KUKA KRL program: PgProg.src

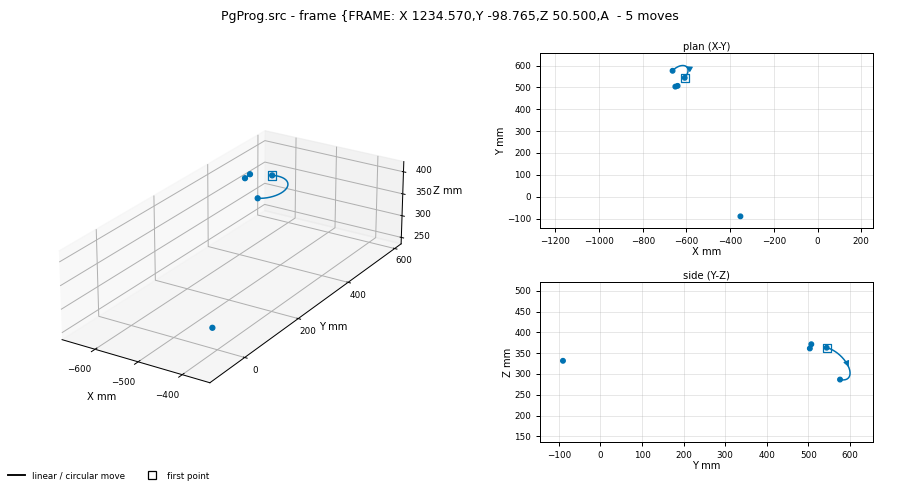
[picture p0: tool path of PgProg.src in frame {FRAME: X 1234.570,Y -98.765,Z 50.500,A , 5 of 9 moves have a stored position in this frame; points joined in program order, loops and branches not executed]
&ACCESS RVP
&REL 1
&PARAM TEMPLATE = C:\KRC\Roboter\Template\vorgabe
&PARAM EDITMASK = *
DEF PgProg ( )


; GLOBAL INTERRUPT DECL 3 WHEN $STOPMESS==TRUE DO IR_STOPM ( )
; INTERRUPT ON 3

;FOLD Initialise and set default speed
BAS (#INITMOV,0)
BAS (#VEL_PTP,100)
BAS (#ACC_PTP,20)
$VEL.CP=0.2
BAS (#TOOL,0)
BAS (#BASE,0)
;ENDFOLD

;;FOLD STARTPOS
;$BWDSTART = FALSE
;PDAT_ACT = PDEFAULT
;BAS(#PTP_DAT)
;FDAT_ACT = {TOOL_NO 0,BASE_NO 0,IPO_FRAME #BASE}
;BAS(#FRAMES)
;;ENDFOLD

$ADVANCE = 5

;FOLD ---- Quickly skip BCO ----
; PTP $AXIS_ACT
;ENDFOLD

;FOLD ---- GO HOME ----
; PTP {A1 0.000, A2 -90.000, A3 90.000, A4 0.000, A5 0.000, A6 0.000, E1 0, E2 0, E3 0, E4 0, E5 0, E6 0}
;ENDFOLD


; Program generated by RoboDK v6.0.7 for KUKA KR 10 R1440-2 on XX/XX/XXXX 18:00:00
; Using nominal kinematics.
; ---- Setting reference (Base) ----
$BASE = {FRAME: X 1234.570,Y -98.765,Z 50.500,A 30.000,B 0.000,C 0.000}
; --------------------------
; ---- Setting tool (TCP) ----
$TOOL = {FRAME: X 10.000,Y 20.000,Z 150.000,A 0.000,B 0.000,C 15.000}
; --------------------------
$VEL.CP = 0.25000
$APO.CPTP = 5
$APO.CDIS = 5.000
PTP {A1 0.00000,A2 -10.00000,A3 20.00000,A4 0.00000,A5 30.00000,A6 0.00000} C_PTP
LIN {X -607.850,Y 543.849,Z 363.215,A 150.000,B 50.000,C -165.000} C_DIS
CIRC {X -602.951,Y 596.788,Z 316.595,A 150.000,B 50.000,C -165.000},{X -663.517,Y 575.988,Z 286.611,A 150.000,B 50.000,C -165.000} C_DIS
PTP {A1 20.00000,A2 -10.00000,A3 20.00000,A4 0.00000,A5 30.00000,A6 0.00000} C_PTP
$ACC.ORI1 = 120.00000
$ACC.ORI2 = 120.00000
$VEL.ORI1 = 60.00000
$VEL.ORI2 = 60.00000
$ACC.CP = 0.80000
$VEL.CP = 0.10000
LIN {X -650.861,Y 503.437,Z 361.399,A 150.000,B 50.000,C -165.000} C_DIS
$APO.CPTP = 0
$APO.CDIS = 0.000
LIN {X -640.584,Y 506.980,Z 371.534,A 150.000,B 50.000,C -165.000} C_DIS
WAIT SEC 0.500
HALT
Wait for StrClear($LOOP_MSG[])
$LOOP_CONT = TRUE
$LOOP_MSG[] = "Hello from postgen"
; a comment
SubProgram()
CustomCode(42)
ThreadProg
$OUT[1]=TRUE
Valve=FALSE
$ANOUT[3]=2.5
WAIT FOR ($IN[2]==TRUE)
START_TIMER:
$TIMER_STOP[1]=TRUE
$TIMER_FLAG[1]=FALSE
$TIMER[1]=1.500
$TIMER_STOP[1]=FALSE
WAIT FOR ($IN[4]==FALSE OR $TIMER_FLAG[1])
$TIMER_STOP[1]=TRUE
IF $TIMER_FLAG[1]== TRUE THEN
    HALT ; Timed out!
    GOTO START_TIMER
ENDIF
; ---- Setting tool (TCP) ----
$TOOL = {FRAME: X 0.000,Y 0.000,Z 200.000,A 0.000,B 0.000,C 0.000}
; --------------------------
PTP {A1 0.00000,A2 -10.00000,A3 20.00000,A4 0.00000,A5 30.00000,A6 0.00000} C_PTP
PTP {A1 10.00000,A2 -5.00000,A3 25.00000,A4 5.00000,A5 35.00000,A6 5.00000} C_PTP
LIN {X -353.026,Y -90.135,Z 331.702,A 178.023,B 40.650,C -169.444} C_DIS
END
